// TIA Portal project "OTOMATIK TRANSFER ASANSORU UYGULAMASI" (V18)

(* hardware
DEVICE "S7-1200 station_1"  S7-1200 Station
   slot 0: "Rack_0"  S7-1200 Rack  Rack  V1.0
   slot 1: "PLC_1"  CPU 1214C AC/DC/Rly  6ES7 214-1BG40-0XB0  V4.6
*)

// ===== PLC "PLC_1"  CPU 1214C AC/DC/Rly =====

VAR_GLOBAL   // PLC tag table "Default tag table"
   "START BUT" AT %I0.0 : Bool;
   "STOP BUT" AT %I0.1 : Bool;
   "ALT PIS GERI SEN" AT %I0.2 : Bool;
   "ALT PIS ILERI SEN" AT %I0.3 : Bool;
   "UST PIS GERI SEN" AT %I0.4 : Bool;
   "UST PIS ILERI SEN" AT %I0.5 : Bool;
   "ASAN ASAGI SEN" AT %I0.6 : Bool;
   "ASAN YUKARI SEN" AT %I0.7 : Bool;
   "URUN TESPIT SEN" AT %I1.0 : Bool;
   "ALT VALF ILERI" AT %Q0.0 : Bool;
   "UST VALF ILERI" AT %Q0.1 : Bool;
   "ASAN VALF YUKARI" AT %Q0.2 : Bool;
   "ASAN VALF  ASAGI" AT %Q0.3 : Bool;
   "GENEL START MEM" AT %M10.0 : Bool;
   "M1" AT %M10.1 : Bool;
   "M2" AT %M10.2 : Bool;
END_VAR

ORGANIZATION_BLOCK "Main"   // OB1, LAD, ProgramCycle
TITLE = "Main Program Sweep (Cycle)"
{ S7_Optimized_Access := 'TRUE' }
VERSION : 0.1
   VAR_INPUT
      Initial_Call : Bool;   // Initial call of this OB
      Remanence : Bool;   // =True, if remanent data are available
   END_VAR
BEGIN

REGION Network 1: SISTEM GENEL START
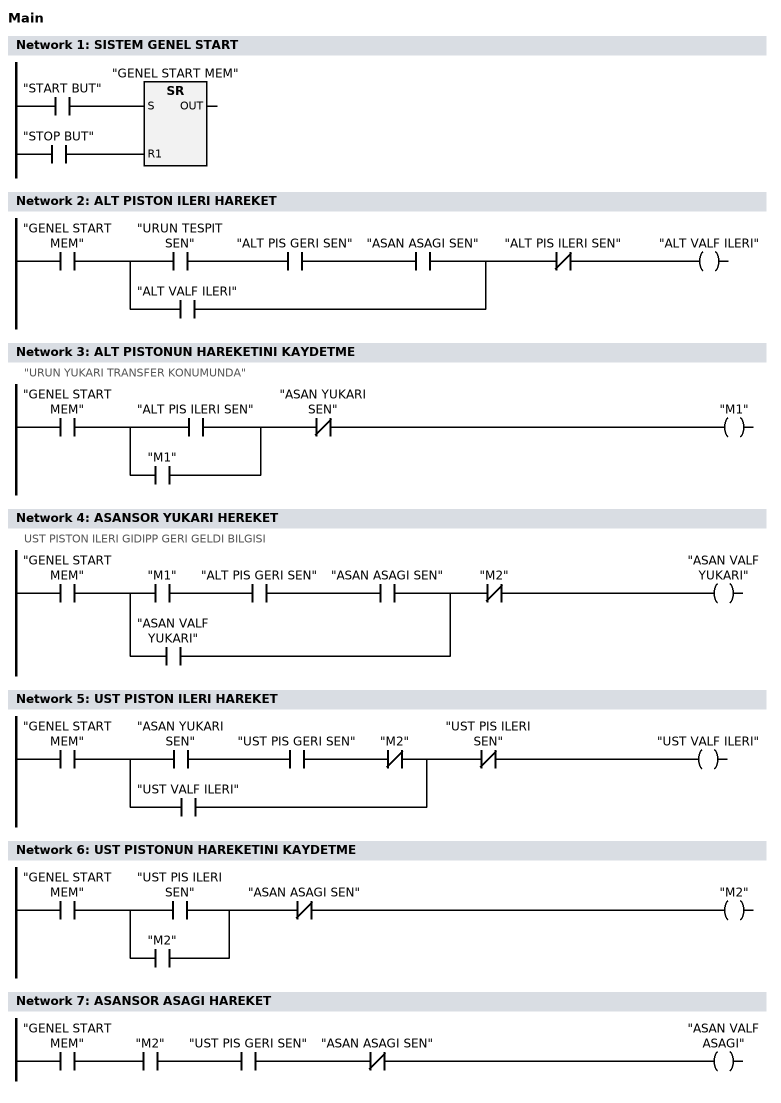
   RUNG wire#powerrail
      Contact( "START BUT" )
      S_SR(operand := "GENEL START MEM", r1 := wire#w1)
   END_RUNG
   RUNG wire#powerrail
      Contact( "STOP BUT" )
   END_RUNG wire#w1
   // the same network as SCL:
   IF "START BUT" THEN
       "GENEL START MEM" := TRUE;   // SR flip-flop
   END_IF;
   IF "STOP BUT" THEN "GENEL START MEM" := FALSE; END_IF;
END_REGION

REGION Network 2: ALT PISTON ILERI HAREKET
   RUNG wire#powerrail
      Contact( "GENEL START MEM" )
      wire#w1
      Contact( "URUN TESPIT SEN" )
      Contact( "ALT PIS GERI SEN" )
      Contact( "ASAN ASAGI SEN" )
      wire#w2
      I_Contact( "ALT PIS ILERI SEN" )
      Coil( "ALT VALF ILERI" )
   END_RUNG
   RUNG wire#w1
      Contact( "ALT VALF ILERI" )
   END_RUNG wire#w2
   // the same network as SCL:
   "ALT VALF ILERI" := "GENEL START MEM" AND (("URUN TESPIT SEN" AND "ALT PIS GERI SEN" AND "ASAN ASAGI SEN") OR "ALT VALF ILERI") AND NOT "ALT PIS ILERI SEN";
END_REGION

REGION Network 3: ALT PISTONUN HAREKETINI KAYDETME
   // "URUN YUKARI TRANSFER KONUMUNDA"
   RUNG wire#powerrail
      Contact( "GENEL START MEM" )
      wire#w1
      Contact( "ALT PIS ILERI SEN" )
      wire#w2
      I_Contact( "ASAN YUKARI SEN" )
      Coil( "M1" )
   END_RUNG
   RUNG wire#w1
      Contact( "M1" )
   END_RUNG wire#w2
   // the same network as SCL:
   "M1" := "GENEL START MEM" AND ("ALT PIS ILERI SEN" OR "M1") AND NOT "ASAN YUKARI SEN";
END_REGION

REGION Network 4: ASANSOR YUKARI HEREKET
   // UST PISTON ILERI GIDIPP GERI GELDI BILGISI
   RUNG wire#powerrail
      Contact( "GENEL START MEM" )
      wire#w1
      Contact( "M1" )
      Contact( "ALT PIS GERI SEN" )
      Contact( "ASAN ASAGI SEN" )
      wire#w2
      I_Contact( "M2" )
      Coil( "ASAN VALF YUKARI" )
   END_RUNG
   RUNG wire#w1
      Contact( "ASAN VALF YUKARI" )
   END_RUNG wire#w2
   // the same network as SCL:
   "ASAN VALF YUKARI" := "GENEL START MEM" AND (("M1" AND "ALT PIS GERI SEN" AND "ASAN ASAGI SEN") OR "ASAN VALF YUKARI") AND NOT "M2";
END_REGION

REGION Network 5: UST PISTON ILERI HAREKET
   RUNG wire#powerrail
      Contact( "GENEL START MEM" )
      wire#w1
      Contact( "ASAN YUKARI SEN" )
      Contact( "UST PIS GERI SEN" )
      I_Contact( "M2" )
      wire#w2
      I_Contact( "UST PIS ILERI SEN" )
      Coil( "UST VALF ILERI" )
   END_RUNG
   RUNG wire#w1
      Contact( "UST VALF ILERI" )
   END_RUNG wire#w2
   // the same network as SCL:
   "UST VALF ILERI" := "GENEL START MEM" AND (("ASAN YUKARI SEN" AND "UST PIS GERI SEN" AND NOT "M2") OR "UST VALF ILERI") AND NOT "UST PIS ILERI SEN";
END_REGION

REGION Network 6: UST PISTONUN HAREKETINI KAYDETME
   RUNG wire#powerrail
      Contact( "GENEL START MEM" )
      wire#w1
      Contact( "UST PIS ILERI SEN" )
      wire#w2
      I_Contact( "ASAN ASAGI SEN" )
      Coil( "M2" )
   END_RUNG
   RUNG wire#w1
      Contact( "M2" )
   END_RUNG wire#w2
   // the same network as SCL:
   "M2" := "GENEL START MEM" AND ("UST PIS ILERI SEN" OR "M2") AND NOT "ASAN ASAGI SEN";
END_REGION

REGION Network 7: ASANSOR ASAGI HAREKET
   RUNG wire#powerrail
      Contact( "GENEL START MEM" )
      Contact( "M2" )
      Contact( "UST PIS GERI SEN" )
      I_Contact( "ASAN ASAGI SEN" )
      Coil( "ASAN VALF  ASAGI" )
   END_RUNG
   // the same network as SCL:
   "ASAN VALF  ASAGI" := "GENEL START MEM" AND "M2" AND "UST PIS GERI SEN" AND NOT "ASAN ASAGI SEN";
END_REGION
END_ORGANIZATION_BLOCK